# B&R Automation Studio project lab2_2 (part 2)

#### gmcipesm.cnc
```
Root (LangModule=ailgcode, Version=1.0)
  AILHeader = def ip_global BOOL  __CANCEL_RND 
    def ip_global BOOL  __C2_SPLINE_ACTIVE 
    def ip_global LREAL __RNDM_RADIUS 
    def ip_global LREAL __CSPLINE_CHORD_ERROR 
    def ip_global DINT __SET_GXX_ACTIVE 
    def ip_global DINT __SET_GXX_REACTIVATE 
    def ip_global DINT __SET_GXX_CALL_CNT 
    def ip_global REAL __VAR1 
    def ip_global DINT __ACTIVE_MIRROR 

    sub OnProgStartPrivate
      %__CANCEL_RND = 0;
      %__RNDM_RADIUS = 0.0;
      %__C2_SPLINE_ACTIVE = 0;
      %__CSPLINE_CHORD_ERROR = 0.001;
      %__SET_GXX_ACTIVE = 0;
      %__SET_GXX_REACTIVATE = 0;
      %__SET_GXX_CALL_CNT = 0;
      %__ACTIVE_MIRROR = 20;
    endsub

    sub EndSplineSection
      
      if (%__C2_SPLINE_ACTIVE)
        `T:GCodes,G802`(:"bc_par":1 :);
        %__C2_SPLINE_ACTIVE = 0;
        
        DispatchMPList(::);
      endif
    endsub
    sub WriteZpTable
      
      #next_motion.Command = MPCMD_SET_ZP_TABLE;
      #next_motion.Data.SetZeroPtTable.ZpRecIdx = $[1];
      #next_motion.Data.SetZeroPtTable.ZpOffset[0] = $[2];
      #next_motion.Data.SetZeroPtTable.ZpOffset[1] = $[3];
      #next_motion.Data.SetZeroPtTable.ZpOffset[2] = $[4];
      PushPacket(::);
      DispatchMPList(::);
    endsub

    sub ReactivateGxx
      
      
      if (%__SET_GXX_CALL_CNT != 0)
          if (%__SET_GXX_REACTIVATE == 1)
            `T:GCodes,G54`(::);
             DispatchMPList(::);
             #sys_vars.ZP = %__SET_GXX_REACTIVATE;
          elif (%__SET_GXX_REACTIVATE == 2)
            `T:GCodes,G55`(::);
             DispatchMPList(::);
             #sys_vars.ZP = %__SET_GXX_REACTIVATE;
          elif (%__SET_GXX_REACTIVATE == 3)
            `T:GCodes,G56`(::);
             DispatchMPList(::);
             #sys_vars.ZP = %__SET_GXX_REACTIVATE;
          elif (%__SET_GXX_REACTIVATE == 4)
            `T:GCodes,G57`(::);
             DispatchMPList(::);
             #sys_vars.ZP = %__SET_GXX_REACTIVATE;
          elif (%__SET_GXX_REACTIVATE == 5)
            `T:GCodes,G58`(::);
             DispatchMPList(::);
             #sys_vars.ZP = %__SET_GXX_REACTIVATE;
          elif (%__SET_GXX_REACTIVATE == 6)
            `T:GCodes,G59`(::);
             DispatchMPList(::);
             #sys_vars.ZP = %__SET_GXX_REACTIVATE;
          endif
          %__SET_GXX_REACTIVATE = 0;
          %__SET_GXX_CALL_CNT = 0;
      endif
    endsub (Append=Yes)
  BuiltInProcs:
    RESET_G54 = WriteZpTable(:1, 0.0, 0.0, 0.0:); (MinArgs=0, MaxArgs=0)
    RESET_G55 = WriteZpTable(:2, 0.0, 0.0, 0.0:); (MinArgs=0, MaxArgs=0)
    RESET_G56 = WriteZpTable(:3, 0.0, 0.0, 0.0:); (MinArgs=0, MaxArgs=0)
    RESET_G57 = WriteZpTable(:4, 0.0, 0.0, 0.0:); (MinArgs=0, MaxArgs=0)
    RESET_G58 = WriteZpTable(:5, 0.0, 0.0, 0.0:); (MinArgs=0, MaxArgs=0)
    RESET_G59 = WriteZpTable(:6, 0.0, 0.0, 0.0:); (MinArgs=0, MaxArgs=0)
    SET_G54 = WriteZpTable(:1, $[1], $[2], $[3]:);
      %_CNC.move_cmd_mode = MPCMD_LIN_INTPOL;
      %__SET_GXX_ACTIVE = 1;
      %__SET_GXX_REACTIVATE = 0;
      %__SET_GXX_CALL_CNT = 0;		
      
      `T:GCodes,G54`(::);
      #sys_vars.ZP = 1; (MinArgs=3, MaxArgs=3)
    SET_G55 = WriteZpTable(:2, $[1], $[2], $[3]:);
      %_CNC.move_cmd_mode = MPCMD_LIN_INTPOL;
      %__SET_GXX_ACTIVE = 2;
      %__SET_GXX_REACTIVATE = 0;
      %__SET_GXX_CALL_CNT = 0;		
      `T:GCodes,G55`(::);
      #sys_vars.ZP = 2; (MinArgs=3, MaxArgs=3)
    SET_G56 = WriteZpTable(:3, $[1], $[2], $[3]:);
      %_CNC.move_cmd_mode = MPCMD_LIN_INTPOL;
      %__SET_GXX_ACTIVE = 3;
      %__SET_GXX_REACTIVATE = 0;
      %__SET_GXX_CALL_CNT = 0;		
      `T:GCodes,G56`(::);
      #sys_vars.ZP = 3; (MinArgs=3, MaxArgs=3)
    SET_G57 = WriteZpTable(:4, $[1], $[2], $[3]:);
      %_CNC.move_cmd_mode = MPCMD_LIN_INTPOL;
      %__SET_GXX_ACTIVE = 4;
      %__SET_GXX_REACTIVATE = 0;
      %__SET_GXX_CALL_CNT = 0;		
      `T:GCodes,G57`(::);
      #sys_vars.ZP = 4; (MinArgs=3, MaxArgs=3)
    SET_G58 = WriteZpTable(:5, $[1], $[2], $[3]:);
      %_CNC.move_cmd_mode = MPCMD_LIN_INTPOL;
      %__SET_GXX_ACTIVE = 5;
      %__SET_GXX_REACTIVATE = 0;
      %__SET_GXX_CALL_CNT = 0;		
      `T:GCodes,G58`(::);
      #sys_vars.ZP = 5; (MinArgs=3, MaxArgs=3)
    SET_G59 = WriteZpTable(:6, $[1], $[2], $[3]:);
      %_CNC.move_cmd_mode = MPCMD_LIN_INTPOL;
      %__SET_GXX_ACTIVE = 6;
      %__SET_GXX_REACTIVATE = 0;
      %__SET_GXX_CALL_CNT = 0;		
      `T:GCodes,G59`(::);
      #sys_vars.ZP = 6; (MinArgs=3, MaxArgs=3)
    RESET_MIRROR = `T:GCodes,G20`(::); (MinArgs=0, MaxArgs=0)
  PVMacros:
    WORKFRAME $WFRAME (ArrayDims=0)
      SET = `T:BuiltInProcs,RESET_SCALING`(::);
        #next_motion.Data.Frame.Data = ${EXPR};
        #next_motion.Command = MPCMD_W_FRAME;
        PushPacket(::); (Inline=Yes)
    WORKFRAME_ADD $WFRAME_ADD (ArrayDims=0)
      SET = `T:BuiltInProcs,RESET_SCALING`(::);
        #next_motion.Data.Frame.Data = ${EXPR};
        #next_motion.Command = MPCMD_W_FRAME_ADD;
        PushPacket(::); (Inline=Yes)
  GCodes:
    G_INIT_ESM = ReactivateGxx(::); (GNum=-5, AutoPush=Yes, Eval=First, Inline=No, GenerateIfGroups=1,1000)
    G_MODAL (GNum=-1, AutoPush=Yes, Group=1000, Eval=Normal, IgnoreIfNoArgs=Yes)
      Arg (ref=dest, MinCount=0, MaxCount=NumAxes, NameType=AXISREF, DataType=PositionValue, WriteOpts=#:u?)
      Arg (ref=center, MinCount=0, MaxCount=3, NameType=InterpolParam, DataType=PositionValue, WriteOpts=#:u?)
      Arg (ref=circlept, MinCount=0, MaxCount=3, NameType=CirclePointParam, DataType=PositionValue, WriteOpts=#:u?)
      Arg (ref=angle, MinCount=0, MaxCount=1, NameType=RotationAngleSpecifier, DataType=RotationAngle, WriteOpts=#:u?)
      Arg (ref=radius, MinCount=0, MaxCount=1, NameType=RadiusSpecifier, DataType=RadiusValue, WriteOpts=#:u?)
    G00 = %_CNC.move_cmd_mode = MPCMD_RAPID_MOVE_INTPOL;
      #sys_vars.modal_grp1_set = 1;
      EndSplineSection(::); (GNum=0, Group=1,50, Inline=Yes, Eval=Early)
    G01 = %_CNC.move_cmd_mode = MPCMD_LIN_INTPOL;
      #sys_vars.modal_grp1_set = 1;
      EndSplineSection(::); (GNum=1, Group=1,50, Inline=Yes, Eval=Early)
    G02 = %_CNC.move_cmd_mode = MPCMD_CIRC_INTPOL_CW;
      #sys_vars.modal_grp1_set = 1;
      EndSplineSection(::); (GNum=2, Group=1,51, Inline=Yes, Eval=Early)
    G03 = %_CNC.move_cmd_mode = MPCMD_CIRC_INTPOL_CCW;
      #sys_vars.modal_grp1_set = 1;
      EndSplineSection(::); (GNum=3, Group=1,51, Inline=Yes, Eval=Early)
    G20 = #next_motion.Command = MPCMD_MIRRORING;
      #next_motion.Data.I4_value = 20;
      %__ACTIVE_MIRROR = #next_motion.Data.I4_value;
      PushPacket(::); (GNum=20, Group=3)
    G20.1 (GNum=20.1, Alias=MIRROR, Group=3)
      Arg (DataType=AXISREF, ref=axis1, MinCount=0, MaxCount=1)
      Arg (DataType=EqString, ref=eq, MinCount=0, MaxCount=1)
      Arg (DataType=FLOAT, ref=dummy_pos1, MinCount=0, MaxCount=1)
      Arg (DataType=AXISREF, ref=axis2, MinCount=0, MaxCount=1)
      Arg (DataType=EqString, ref=eq, MinCount=0, MaxCount=1)
      Arg (DataType=FLOAT, ref=dummy_pos2, MinCount=0, MaxCount=1)
    G20.2 (GNum=20.2, Alias=AMIRROR, Group=3)
      Arg (DataType=AXISREF, ref=axis1, MinCount=1, MaxCount=1)
      Arg (DataType=EqString, ref=eq, MinCount=0, MaxCount=1)
      Arg (DataType=FLOAT, ref=dummy_pos1, MinCount=0, MaxCount=1)
      Arg (DataType=AXISREF, ref=axis2, MinCount=0, MaxCount=1)
      Arg (DataType=EqString, ref=eq, MinCount=0, MaxCount=1)
      Arg (DataType=FLOAT, ref=dummy_pos2, MinCount=0, MaxCount=1)
    G21 = #next_motion.Command = MPCMD_MIRRORING;
      #next_motion.Data.I4_value = 21;
      %__ACTIVE_MIRROR = #next_motion.Data.I4_value;
      PushPacket(::); (GNum=21, Group=3)
    G22 = #next_motion.Command = MPCMD_MIRRORING;
      #next_motion.Data.I4_value = 22;
      %__ACTIVE_MIRROR = #next_motion.Data.I4_value;
      PushPacket(::); (GNum=22, Group=3)
    G23 = #next_motion.Command = MPCMD_MIRRORING;
      #next_motion.Data.I4_value = 23;
      %__ACTIVE_MIRROR = #next_motion.Data.I4_value;
      PushPacket(::); (GNum=23, Group=3)
    G25.1 (GNum=25.1, Group=11, Alias=RNDM)
      Arg (NameType=EqString, DataType=TangArcRadius, ref=radius)
    G25.2 (GNum=25.2, Group=11, Alias=RND)
      Arg (NameType=EqString, DataType=TangArcRadius, ref=radius)
    G53 = #next_motion.Command = MPCMD_ABS_ZP_SHIFT;
      #next_motion.Data.AbsZeroPtShift.ZpRecIdx = 0;
      PushPacket(::);
      #sys_vars.ZP = 0;
      
      %__SET_GXX_REACTIVATE = %__SET_GXX_ACTIVE;
      %__SET_GXX_CALL_CNT = 0; (GNum=53, Group=6, AllowGroups=8,19,21,100,101,102,103)
    G92 (GNum=92, Group=21, ResetArgs=Yes, AllowGroups=6,8,19,32,100,101,102,103)
      Arg (NameType=AXISREF, DataType=PositionValue, ref=offset, MinCount=0, MaxCount=NumAxes, WriteOpts=#:u?)
      Arg (NameType=RotationAngleSpecifier, DataType=RotationAngle, ref=h_rot, MinCount=0, MaxCount=1, WriteOpts=#:u?, DenyArgs=3,4,5)
      Arg (NameType=EulerAngleName, DataType=RotationAngle, ref=e_rot, MinCount=0, MaxCount=3, WriteOpts=#:u?, DenyArgs=2,4,5)
      Arg (NameType=RPYAngleName, DataType=RotationAngle, ref=rpy_rot, MinCount=0, MaxCount=3, WriteOpts=#:u?, DenyArgs=2,3,5)
      Arg (NameType=RotaryVectorName, DataType=RotaryVector, ref=matrix, MinCount=0, MaxCount=3, WriteOpts=#:u?, DenyArgs=2,3,4)
    G92.1 (GNum=92.1, Group=21, ALIAS=SCALE, AliasIsPattern=Yes)
      Arg (DataType=FLOAT, ref=factor, MinCount=0, MaxCount=1)
    G92.2 (GNum=92.2, Group=21, ALIAS=ASCALE, AliasIsPattern=Yes)
      Arg (DataType=FLOAT, ref=factor, MinCount=1, MaxCount=1)
    G492 (GNum=492, Group=490, Alias=TRANS, AllowGroups=9999)
      Arg (NameType=AXISREF, DataType=PositionValue, ref=offsets, MinCount=0, MaxCount=NumAxes, WriteOpts=#:)
    G494 (GNum=494, Group=490, Alias=ROT, AllowGroups=9999, MinArgs=0, MaxArgs=1)
      Arg RPLArgPrefix (DataType=FLOAT, ref=rpl_value, MinCount=0, MaxCount=1, DenyArgs=offsets)
      Arg (NameType=AXISREF, DataType=PositionValue, ref=offsets, MinCount=0, MaxCount=NumAxes, DenyArgs=rpl_value, WriteOpts=#:)
    G500 = %__SET_GXX_REACTIVATE = 0;
       %__SET_GXX_ACTIVE = 0;
       %__SET_GXX_CALL_CNT = 0;
      `T:GCodes,G53`(::); (GNum=500, Group=6, AllowGroups=8,19,21,100,101,102,103)
    G804 = if (!%__C2_SPLINE_ACTIVE)
         
        `T:GCodes,G801`(:"seg_type":"CE", "seg_par":%__CSPLINE_CHORD_ERROR, "bc_par":1 :);
        %__C2_SPLINE_ACTIVE = 1;
        
        DispatchMPList(::);
        
        %_CNC.move_cmd_mode = MPCMD_LIN_INTPOL;
      endif (GNum=804, Alias=CSPLINE)
```

### Data object Logical/GmcIpConfig/gmcipmxd (Cnc, version 5.02.1)

#### gmcipmxd.cnc
```
(********************************************************************
 * COPYRIGHT (C) B&R Industrial Automation GmbH
 ********************************************************************
 * Library: Motion Command Extension
 * File: arnc0mx.typ
 * Author: B&R
 ********************************************************************
 * Data types of Motion Command Library
 ********************************************************************)

TYPE
	MXOrientationType : STRUCT
		Type : UDINT;
		Angle : ARRAY[0..3]OF LREAL;
	END_STRUCT;
	MXPositionType : STRUCT
		x : LREAL;
		y : LREAL;
		z : LREAL;
	END_STRUCT;
	MXFrameType : 	STRUCT
		Pos : MXPositionType;
		Orient : MXOrientationType;
	END_STRUCT;
	MXToolType : STRUCT
		Index : UDINT;
		Frame : MXFrameType;
		Radius : LREAL;
	END_STRUCT;
	MXJointAxisType :ARRAY[0..5]OF LREAL;
	MXAuxAxisType :ARRAY[0..14]OF LREAL;
	MXBaseAxisType :ARRAY[0..5]OF LREAL;
	MXRotAxisType :ARRAY[0..5]OF LREAL;
	MXConfigType : 	STRUCT
		Mode : UDINT;
	END_STRUCT;
	MXPointType : 	STRUCT
		Pos : MXPositionType;
		Orient : MXOrientationType;
		Cfg : MXConfigType;
		RotAxis : MXRotAxisType;
		AuxAxis : MXAuxAxisType;
	END_STRUCT;
	MXPathTransType : STRUCT
		Radius	:	LREAL;
		Type	:	UDINT;
	END_STRUCT;
	MXPathDescType : STRUCT
		Trans	:	MXPathTransType;
	END_STRUCT;
	MXOptMotType : STRUCT
		Enable : BOOL;
		VelPathDef : USINT;
		RobotPar : USINT;
		Limits : USINT;
	END_STRUCT;
	MXDynamicDescType :	STRUCT
		Accel : LREAL := 100;
		Decel : LREAL := 100;
		Optmot : MXOptMotType;
	END_STRUCT;
	MXHWTrigType : 	STRUCT
		Source : USINT;
		Index : USINT;
	END_STRUCT;
	MXSWTrigType : STRUCT
		Expression : STRING[64];
	END_STRUCT;
	MXTriggConfigType :	STRUCT
		Type : UINT;
		HWTrig : MXHWTrigType;
		SWTrig : MXSWTrigType;
		Edge : USINT;
		ResidPath : USINT;
	END_STRUCT;
	MXVelocityType : STRUCT
		v : LREAL;
		Mode : UDINT := 1;
	END_STRUCT;
	MXAxisTargetType : 	STRUCT
		JointAxis : MXJointAxisType;
		AuxAxis : MXAuxAxisType;
		BaseAxis : MXBaseAxisType;
	END_STRUCT;
	MXCDCType : STRUCT
		ArcTransSpd : LREAL := 100;
		SpdMode : UDINT;
		ContourViolation : UDINT;
		TransMode : UDINT;
		EntryMode : USINT;
		AcrToLine : BOOL;
	END_STRUCT;
	MXAutoTangType : STRUCT
		Offset : LREAL;
	END_STRUCT;
	MXHWTriggerType :	STRUCT
		Source : UINT;
		Index : UINT;
	END_STRUCT;
	MXTriggerConfigType : 	STRUCT
		Type : UINT;
		Edge : UINT;
		HWTrigger : MXHWTriggerType;
	END_STRUCT;
END_TYPE

(********************************************************************
 * COPYRIGHT (C) B&R Industrial Automation GmbH
 ********************************************************************
 * Library: ARNC0MX
 * File: arnc0mx.fun
 * Created: 13.06.2012
 ********************************************************************
 * Functions and function blocks of library ARNC0MX
 ********************************************************************)
FUNCTION MXPointToJointEx1 : UDINT
	VAR_INPUT
		AddrTrfData : UDINT;
		Point : MXPointType;
		Joint : MXJointAxisType;
		TrfType : UDINT;
		Tool : MXToolType;
		BaseFrame : MXFrameType;
		RefJoint : ARRAY[0..5] OF LREAL;
	END_VAR
END_FUNCTION

FUNCTION MXPointToJointEx : UDINT
	VAR_INPUT
		AddrTrfData : UDINT;
		Point : MXPointType;
		Joint : MXJointAxisType;
		TrfType : UDINT;
		Tool : MXToolType;
		BaseFrame : MXFrameType;
		RefJoint : MXJointAxisType;
	END_VAR
END_FUNCTION

FUNCTION MXJointToPointEx1 : UDINT
	VAR_INPUT
		AddrTrfData : UDINT;
		Joint : MXJointAxisType;
		Point : MXPointType;
		AnglesType : UDINT;
		TrfType : UDINT;
		Tool : MXToolType;
		BaseFrame : MXFrameType;
		RefPath : ARRAY[0..5] OF LREAL;
	END_VAR
END_FUNCTION

FUNCTION MXJointToPointEx : UDINT
	VAR_INPUT
		AddrTrfData : UDINT;
		Joint : MXJointAxisType;
		Point : MXPointType;
		AnglesType : UDINT;
		TrfType : UDINT;
		Tool : MXToolType;
		BaseFrame : MXFrameType;
		RefPoint : MXPointType;
	END_VAR
END_FUNCTION

FUNCTION MXCncAxesToPoint : UDINT
	VAR_INPUT
		AddrTrfData : UDINT;
		Axis : ARRAY[0..14] OF LREAL;
		Point : MXPointType;
		TrfType : UDINT;
		AnglesType : UDINT;
		AxisMapCode : ARRAY[0..14] OF UINT;
		AxisMapIdx : ARRAY[0..14] OF UINT;
		ActiveAxesCount : UDINT;
	END_VAR
END_FUNCTION

FUNCTION MXFromOrient : UDINT
	VAR_INPUT
		Orient : MXOrientationType;
		Matrix : ARRAY[0..8] OF LREAL;
	END_VAR
END_FUNCTION

FUNCTION MXToOrient : UDINT
	VAR_INPUT
		Matrix : ARRAY[0..8] OF LREAL;
		Type : UDINT;
		Orient : MXOrientationType;
		RefAngle : ARRAY[0..2] OF LREAL;
	END_VAR
END_FUNCTION

FUNCTION MXConvertOrient : UDINT
	VAR_INPUT
		OrientIn : MXOrientationType;
		Type : UDINT;
		OrientOut : MXOrientationType;
		RefAngle : ARRAY[0..2] OF LREAL;
	END_VAR
END_FUNCTION

FUNCTION MXFrameRotX : UDINT
	VAR_INPUT
		Frame : MXFrameType;
		Angle : LREAL;
	END_VAR
END_FUNCTION

FUNCTION MXFrameRotY : UDINT
	VAR_INPUT
		Frame : MXFrameType;
		Angle : LREAL;
	END_VAR
END_FUNCTION

FUNCTION MXFrameRotZ : UDINT
	VAR_INPUT
		Frame : MXFrameType;
		Angle : LREAL;
	END_VAR
END_FUNCTION

FUNCTION MXFrameEuler : UDINT
	VAR_INPUT
		Frame : MXFrameType;
		Phi : LREAL;
		Theta : LREAL;
		Psi : LREAL;
	END_VAR
END_FUNCTION

FUNCTION MXFrameRPY : UDINT
	VAR_INPUT
		Frame : MXFrameType;
		Roll : LREAL;
		Pitch : LREAL;
		Yaw : LREAL;
	END_VAR
END_FUNCTION

FUNCTION MXFrameTrans : UDINT
	VAR_INPUT
		Frame : MXFrameType;
		DistanceX : LREAL;
		DistanceY : LREAL;
		DistanceZ : LREAL;
	END_VAR
END_FUNCTION

FUNCTION MXFrameTransX : UDINT
	VAR_INPUT
		Frame : MXFrameType;
		Distance : LREAL;
	END_VAR
END_FUNCTION

FUNCTION MXFrameTransY : UDINT
	VAR_INPUT
		Frame : MXFrameType;
		Distance : LREAL;
	END_VAR
END_FUNCTION

FUNCTION MXFrameTransZ : UDINT
	VAR_INPUT
		Frame : MXFrameType;
		Distance : LREAL;
	END_VAR
END_FUNCTION

FUNCTION MXFrameApply : UDINT
	VAR_INPUT
		Frame1 : MXFrameType;
		Frame2 : MXFrameType;
	END_VAR
END_FUNCTION

FUNCTION MXFromFrame : UDINT
	VAR_INPUT
		Frame : MXFrameType;
		PointIn : MXPointType;
		PointOut : MXPointType;
	END_VAR
END_FUNCTION

FUNCTION MXToFrame : UDINT
	VAR_INPUT
		Frame : MXFrameType;
		PointIn : MXPointType;
		PointOut : MXPointType;
	END_VAR
END_FUNCTION

(********************************************************************
 * COPYRIGHT (C) B&R Industrial Automation GmbH
 ********************************************************************
 * Library: Motion Command Extension
 * File: arnc0mx.var
 * Author: B&R
 ********************************************************************
 * Constants of Motion Command Library
 ********************************************************************)

(* Velocity mode constants (<MXVelocityType>.Mode) *)
VAR CONSTANT
  MX_VEL_MODE_RAPID : UDINT := 0; (* rapid mode *)
  MX_VEL_MODE_FEED  : UDINT := 1; (* feedrate mode *)
  MX_VEL_MODE_TIME  : UDINT := 2; (* inverse time mode *)
END_VAR

(* MXVelocityType constants *)
VAR CONSTANT
  MX_VEL_RAPID  : MXVelocityType := (Mode:=0);           (* rapid movement         *)
  MX_VEL_F50000 : MXVelocityType := (v:=50000, Mode:=1); (* 50000 units per minute *)
  MX_VEL_F10000 : MXVelocityType := (v:=10000, Mode:=1); (* 10000 units per minute *)
  MX_VEL_F5000  : MXVelocityType := (v:=5000,  Mode:=1); (* 5000 units per minute  *)
  MX_VEL_F1000  : MXVelocityType := (v:=1000,  Mode:=1); (* 1000 units per minute  *)
  MX_VEL_F500   : MXVelocityType := (v:=500,   Mode:=1); (* 500 units per minute   *)
  MX_VEL_F100   : MXVelocityType := (v:=100,   Mode:=1); (* 100 units per minute   *)
END_VAR

(* Trigger configuration constants *)
VAR CONSTANT
  MX_TRIGGER_HW	            : UINT := 0;           (* Hardware trigger - MXHWTriggerType *)
  MX_TRIGGER_POSITIVE_EDGE  : UINT := 0;           (* Positive edge						 *)
  MX_TRIGGER_NEGATIVE_EDGE  : UINT := 1;           (* Negative edge						 *)
  MX_TRIGGER_HW_INPUT1		: UINT := 1;           (* Hardware trigger input 1			 *)
  MX_TRIGGER_HW_INPUT2		: UINT := 2;           (* Hardware trigger input 1			 *)
END_VAR

(* MXFrameMXFrameType constants *)
VAR CONSTANT
  MX_FRM_ZERO : MXFrameType := (0); (* zero (identity) frame *)
END_VAR

(* Transition type constants (<MXPathTransType>.Type) *)
VAR CONSTANT
  MX_TRANS_OFF      : UDINT := 0; (* Transition deactivated *)
  MX_TRANS_ACCURATE : UDINT := 1; (* Accuracy hold *)
  MX_TRANS_ARC      : UDINT := 2; (* Tangential transition arcs *)
  MX_TRANS_ROUND    : UDINT := 3; (* Rounding edges *)
END_VAR

(* Orientation type constants (<MXOrientationType>.Type) matches constants from TRF_LIB *)
VAR CONSTANT
  MX_CARDAN_XYZ_ANGLES    : UDINT := 1;      (* Cardan XYZ angles *)
  MX_EULER_XYZ_ANGLES     : UDINT := 1;      (* Cardan XYZ angles *)
  MX_CARDAN_XZY_ANGLES    : UDINT := 2;      (* Cardan XZY angles *)
  MX_EULER_XZY_ANGLES     : UDINT := 2;      (* Cardan XZY angles *)
  MX_CARDAN_YXZ_ANGLES    : UDINT := 4;      (* Cardan YXZ angles *)
  MX_EULER_YXZ_ANGLES     : UDINT := 4;      (* Cardan YXZ angles *)
  MX_CARDAN_YZX_ANGLES    : UDINT := 8;      (* Cardan YZX angles *)
  MX_EULER_YZX_ANGLES     : UDINT := 8;      (* Cardan YZX angles *)
  MX_CARDAN_ZXY_ANGLES    : UDINT := 16;     (* Cardan ZXY angles *)
  MX_EULER_ZXY_ANGLES     : UDINT := 16;     (* Cardan ZXY angles *)
  MX_CARDAN_ZYX_ANGLES    : UDINT := 32;     (* Cardan ZYX angles *)
  MX_EULER_ZYX_ANGLES     : UDINT := 32;     (* Cardan ZYX angles *)
  MX_EULER_XYX_ANGLES     : UDINT := 64;     (* Euler XYX angles  *)
  MX_EULER_XZX_ANGLES     : UDINT := 128;    (* Euler XZX angles  *)
  MX_EULER_YXY_ANGLES     : UDINT := 256;    (* Euler YXY angles  *)
  MX_EULER_YZY_ANGLES     : UDINT := 512;    (* Euler YZY angles  *)
  MX_EULER_ZXZ_ANGLES     : UDINT := 1024;   (* Euler ZXZ angles  *)
  MX_EULER_ZYZ_ANGLES     : UDINT := 2048;   (* Euler ZYZ angles  *)
  MX_POSITIVE_ANGLES      : UDINT := 4096;   (* mathematically positive angles *)
  MX_NEGATIVE_ANGLES      : UDINT := 8192;   (* mathematically negative angles *)
  MX_DIRECT_ANGLES        : UDINT := 16384;  (* direct "R" rotation matrix     *)
  MX_INDIRECT_ANGLES      : UDINT := 32768;  (* indirect "R^T" rotation matrix *)
  MX_EULER_ANGLES         : UDINT := 1024;   (* Euler ZXZ is commonly in view  *)
  MX_CARDAN_ANGLES        : UDINT := 1;      (* Cardan XYZ is commonly in view *)
  MX_NAUTICAL_ANGLES      : UDINT := 1;      (* Cardan XYZ is commonly in view *)
  MX_TAIT_BRYAN_ANGLES    : UDINT := 1;      (* Cardan XYZ is commonly in view *)
  MX_QUATERNION           : UDINT := 8000;   (* quaternion *)
END_VAR

(* Kinematics configuration mode constants (<MXConfigType>.Mode) matches constants from TRF_LIB *)
VAR CONSTANT
  MX_MODE_FRONT           : UDINT := 1;          (* front *)
  MX_MODE_BACK            : UDINT := 2;          (* back *)
  MX_MODE_CONVEX          : UDINT := 4;          (* convex *)
  MX_MODE_CONCAVE         : UDINT := 8;          (* concave *)
  MX_MODE_POSITIVE        : UDINT := 16;         (* positive *)
  MX_MODE_NEGATIVE        : UDINT := 32;         (* negative *)
  MX_MODE_LEFT            : UDINT := 64;         (* left *)
  MX_MODE_RIGHT           : UDINT := 128;        (* right *)
  MX_MODE_DIRECT          : UDINT := 256;        (* direct *)
  MX_MODE_INDIRECT        : UDINT := 512;        (* indirect *)
  MX_MODE_CONVEX2         : UDINT := 1024;       (* convex2 *)
  MX_MODE_CONCAVE2        : UDINT := 2048;       (* concave2 *)
  MX_MODE_CONVEX3         : UDINT := 4096;       (* convex3 *)
  MX_MODE_CONCAVE3        : UDINT := 8192;       (* concave3 *)
  MX_MODE_HETEROGENEOUS   : UDINT := 16384;      (* heterogeneous *)
  MX_MODE_HOMOGENEOUS     : UDINT := 32768;      (* homogeneous *)
  MX_MODE_LEFT2           : UDINT := 65536;      (* left2 *)
  MX_MODE_RIGHT2          : UDINT := 131072;     (* right2 *)
  MX_MODE_NEG_DIR         : UDINT := 268435456;  (* negative direction forced *)
  MX_MODE_POS_DIR         : UDINT := 536870912;  (* positive direction forced *)
  MX_MODE_IN_SW_ENDS      : UDINT := 1073741824; (* in SW ends *)
END_VAR

(* Cutter diameter compensation constants *)
VAR CONSTANT
  MX_CDC_LEFT                    : UDINT := 0;      (* CDC left *)
  MX_CDC_RIGHT                   : UDINT := 1;      (* CDC right *)
  MX_CDC_SPD_ON_CONTOUR          : UDINT := 0;      (* Path speed moves to the contour *)
  MX_CDC_SPD_ON_TCP              : UDINT := 1;      (* Path speed moves to the center of the tool *)
  MX_CDC_NO_COUNTER_VIOLATION    : UDINT := 0;      (* Do NOT allow contour violations due to very short path *)
  MX_CDC_VIOLATION_SHORT_PATH    : UDINT := 1;      (* Allow contour violations due to very short path sections *)
  MX_CDC_VIOLATION_INNER_EDGE    : UDINT := 2;      (* Allow contour violations due to an inner edge without intersection *)
  MX_CDC_LINEAR_TRANSITION       : UDINT := 0;      (* CDC with linear transitions *)
  MX_CDC_ARC_TRANSITION          : UDINT := 1;      (* CDC with arc transitions *)
  MX_CDC_ENTRY_BLOCK             : UDINT := 0;      (* Activate/deactivate CDC indirectly with transi-tion block *)
  MX_CDC_ENTRY_DIRECT            : UDINT := 1;      (* Activate/deactivate CDC directly *)
  MX_CDC_ENTRY_INDIRECT          : UDINT := 2;      (* Activate/deactivate CDC indirectly *)
  MX_CDC_NO_ARC_TO_LINE          : UDINT := 0;      (* Deactivate replacement of arc with straight line *)
  MX_CDC_ARC_TO_LINE             : UDINT := 1;      (* Activate replacement of arc with straight line *)
END_VAR

(* Transformation function types *)
VAR CONSTANT
  MX_TRF_TYPE_INVERSE            : UDINT := 0;      (* TRF_inverse  function *)
  MX_TRF_TYPE_INVERSE2           : UDINT := 1;      (* TRF_inverse2 function *)
  MX_TRF_TYPE_INVERSE3           : UDINT := 2;      (* TRF_inverse3 function *)
  MX_TRF_TYPE_DIRECT             : UDINT := 0;      (* TRF_direct   function *)
  MX_TRF_TYPE_DIRECT2            : UDINT := 1;      (* TRF_direct2  function *)
  MX_TRF_TYPE_DIRECT3            : UDINT := 2;      (* TRF_direct3  function *)
END_VAR

(* Statuses, warnings, errors *)
VAR CONSTANT
  MX_OK                          : UDINT := 0;     (* Status OK *)
  MX_WARNING_AXES                : UDINT := 2001;  (* Transformation returns valid values with warnings on axes *)
  MX_WARNING_REF_POINT_ANGLES    : UDINT := 2002;  (* Values in reference point or reference joint axes may be ignored due to conversion to another angles type *)
  MX_ERROR_WRONG_ANGLE_TYPE      : UDINT := 6001;  (* Angles type is not supported *)
  MX_ERROR_TRF_DATA_NOT_DEFINED  : UDINT := 6002;  (* Address of the transformation data variable is zero *)
  MX_ERROR_WRONG_ROBOT           : UDINT := 6003;  (* Robot is not supported *)
  MX_ERROR_WRONG_TRF_TYPE        : UDINT := 6004;  (* Transformation type not supported *)
  MX_ERROR_TRF_LIB_NOT_SUPPORTED : UDINT := 6005;  (* Transformation library of not supported version *)
  MX_ERROR_TRF_CMD_CODE			 : UDINT := 8001;  (* Unknown command code *)
  MX_ERROR_TRF_MEASURE           : UDINT := 8002;  (* Unknown measure *)
  MX_ERROR_TRF_ANGLES_TYPE       : UDINT := 8003;  (* Unknown angles type *)
  MX_ERROR_TRF_GEN29_CMD_CODE    : UDINT := 9001;  (* Unknown command code *)
  MX_ERROR_UNKNOWN_ROBOT         : UDINT := 9002;  (* Unknown robot *)
  MX_ERROR_INVALID_TRF_TYPE      : UDINT := 9003;  (* Invalid type of transformation *)
  MX_ERROR_TRF_ERROR_AXES        : UDINT := 10003; (* Transformation function returns error of axis *)
  MX_ERROR_TRF_NOT_LICENSED      : UDINT := 10008; (* Transformation function not licenced *)
  MX_ERROR_TRF_NOT_SUPPORTED     : UDINT := 10009; (* Transformation function not supported *)
  MX_ERROR_FCT_NOT_DEFINED       : UDINT := 10010; (* Transformation function address is zero *)
  MX_ERROR_TRF_INVALID_INPUTS    : UDINT := 10015; (* Invalid inputs for transformation error *)
END_VAR

(* Error offsets *)
VAR CONSTANT
  MX_OFFSET_WARNING              : UDINT := 2000;  (* ARNC0MX warnings *)
  MX_OFFSET_WARNING_TRF_FUN      : UDINT := 4000;  (* TRF_LIB warnings *)
  MX_OFFSET_ERROR                : UDINT := 6000;  (* ARNC0MX errros *)
  MX_OFFSET_ERROR_TRF_FUN        : UDINT := 12000; (* TRF_LIB errors *)
END_VAR

(********************************************************************
 * COPYRIGHT (C) B&R Industrial Automation GmbH
 ********************************************************************
 * Library: Motion Command Library
 * File: arnc0mxsv.var
 * Author: B&R
 ********************************************************************
 * System Variables of Motion Command Library
 ********************************************************************)
VAR {SHARED_IP_GLOBAL}
   _Frm  : MXFrameType;
   _Tool : MXToolType;
   _Vel  : MXVelocityType;
   _Base : MXFrameType;
   _Ref  : MXJointAxisType;
   _Pth  : MXPathDescType;
   _Dyn  : MXDynamicDescType;
END_VAR

VAR CONSTANT
   FRM_0   : MXFrameType := (0);
   POINT_0 : MXPointType := (0);
   BASE_0  : MXFrameType := (0);
   TOOL_0  : MXToolType  := (0);
   VEL_0   : MXVelocityType := (Mode:=1);
   REF_0   : MXJointAxisType := (0);
   VEC6_0  : ARRAY[0..5] OF LREAL := 6(0.0);
   PTH_0   : MXPathDescType := (0);
   DYN_0   : MXDynamicDescType := (Accel:=100, Decel:=100);
   AXIS_TARGET_0 : MXAxisTargetType := (0);
END_VAR

VAR {SHARED_IP_GLOBAL}
  __tmp_point : MXPointType;
  __tmp_frame : MXFrameType;
  __tmp_tool : MXToolType;
  __tmp_vel : MXVelocityType;
  __tmp_joint_axis : MXJointAxisType;
  __tmp_axis_target : MXAxisTargetType;
  __tmp_pth : MXPathDescType;
  __tmp_dynamic : MXDynamicDescType;
  __tmp_cdc : MXCDCType;
  __tmp_auto_tang : MXAutoTangType;
  __tmp_trigger : MXTriggerConfigType;
  __mx_status : UDINT;
  __tmp_vec6 : ARRAY[0..5] OF LREAL;
  __tmp_set_pos : ARRAY[0..14] OF LREAL;
  __tmp_axis_code : ARRAY[0..14] OF UINT;
  __tmp_axis_idx : ARRAY[0..14] OF UINT;
END_VAR
```

### Data object Logical/GmcIpConfig/gmcipmx (Cnc, version 5.02.1)

#### gmcipmx.cnc
```
Root (LangModule=ailgcode, Version=1.0)
  AILHeader = sub OnProgStartPrivate
      %_Frm = %FRM_0;
      %_Base = %BASE_0;
      %_Tool = %TOOL_0;
      %_Vel = %VEL_0;
      %_Pth = %PTH_0;
      %_Dyn = %DYN_0;
      if (%_CNC.optmot_segmentation_on)
        %_Dyn.Optmot.Enable = 1 
      endif      
      BlockCpy(:\%_Ref, \%REF_0:);
    endsub
  BuiltInProcs:
    WAIT_PP_SYNC = #next_motion.Command = MPCMD_IP_SYNCH_PP;
      PushPacket(::);
      DispatchAndWait(:IPCMD_SYNC_PP_CONT:);
    ERROR_EX = ErrorEx(:"id":$[1],"fmt":$[2],"data":(:$[3],$[4],$[5],$[6],$[7],$[8],$[9],$[10],$[11],$[12],$[13],$[14]:):); (MinArgs=3, MaxArgs=14)
    SET_POINT:
      Arg (ref=POINT, DataType=ANY_DATA, MinCount=1, MaxCount=1)
    SET_TRIGGER_CONFIG:
      Arg (ref=TRIGGER, DataType=ANY_DATA, MinCount=1, MaxCount=1)
      Arg (ref=bHALT, DataType=ANY_DATA, MinCount=1, MaxCount=1)
      Arg (ref=ID, DataType=ANY_DATA, MinCount=1, MaxCount=1)
    SET_WANTED_JOINT:
      Arg (ref=Ref, DataType=ANY_DATA, MinCount=1, MaxCount=1)
    SET_CIRCLE:
      Arg (ref=END_POINT, DataType=ANY_DATA, MinCount=1, MaxCount=1)
      Arg (ref=CIRCLE_POINT, DataType=ANY_DATA, MinCount=1, MaxCount=1)
      Arg (ref=Angle, DataType=IEC_LREAL, MinCount=0, MaxCount=1)
    SET_AXIS_TARGET:
      Arg (ref=AXIS_TARGET, DataType=ANY_DATA, MinCount=1, MaxCount=1)
    SET_FRAME:
      Arg (ref=Frm, DataType=ANY_DATA, MinCount=0, MaxCount=1)
    SET_BASEFRAME:
      Arg (ref=Base, DataType=ANY_DATA, MinCount=0, MaxCount=1)
    SET_TOOL:
      Arg (ref=Tool, DataType=ANY_DATA, MinCount=0, MaxCount=1)
    SET_PATH_DESC:
      Arg (ref=Pth, DataType=ANY_DATA, MinCount=0, MaxCount=1)
    SET_DYNAMIC_DESC:
      Arg (ref=Dyn, DataType=ANY_DATA, MinCount=0, MaxCount=1)
    SET_VELOCITY:
      Arg (ref=Vel, DataType=ANY_DATA, MinCount=0, MaxCount=1)
    JointToPoint:
      Arg (ref=Joint, UserType=MXJointAxisType, MinCount=1, MaxCount=1)
      Arg (ref=Point, UserType=MXPointType, MinCount=1, MaxCount=1)
    PointToJoint:
      Arg (ref=Point, UserType=MXPointType, MinCount=1, MaxCount=1)
      Arg (ref=Joint, UserType=MXJointAxisType, MinCount=1, MaxCount=1)
    MoveL:
      Arg (ref=POINT, UserType=MXPointType, MinCount=1, MaxCount=1)
      Arg (ref=Frm, UserType=MXFrameType, MinCount=0, MaxCount=1)
      Arg (ref=Base, UserType=MXFrameType, MinCount=0, MaxCount=1)
      Arg (ref=Tool, UserType=MXToolType, MinCount=0, MaxCount=1)
      Arg (ref=Vel, UserType=MXVelocityType, MinCount=0, MaxCount=1)
      Arg (ref=Pth, UserType=MXPathDescType, MinCount=0, MaxCount=1)
      Arg (ref=Dyn, UserType=MXDynamicDescType, MinCount=0, MaxCount=1)
    MoveJ:
      Arg (ref=POINT, UserType=MXPointType, MinCount=1, MaxCount=1)
      Arg (ref=Frm, UserType=MXFrameType, MinCount=0, MaxCount=1)
      Arg (ref=Base, UserType=MXFrameType, MinCount=0, MaxCount=1)
      Arg (ref=Tool, UserType=MXToolType, MinCount=0, MaxCount=1)
      Arg (ref=Vel, UserType=MXVelocityType, MinCount=0, MaxCount=1)
      Arg (ref=Ref, UserType=MXJointAxisType, MinCount=0, MaxCount=1)
      Arg (ref=Pth, UserType=MXPathDescType, MinCount=0, MaxCount=1)
      Arg (ref=Dyn, UserType=MXDynamicDescType, MinCount=0, MaxCount=1)
    MoveC:
      Arg (ref=END_POINT, UserType=MXPointType, MinCount=1, MaxCount=1)
      Arg (ref=CIRCLE_POINT, UserType=MXPointType, MinCount=1, MaxCount=1)
      Arg (ref=Angle, DataType=IEC_LREAL, MinCount=0, MaxCount=1)
      Arg (ref=Frm, UserType=MXFrameType, MinCount=0, MaxCount=1)
      Arg (ref=Base, UserType=MXFrameType, MinCount=0, MaxCount=1)
      Arg (ref=Tool, UserType=MXToolType, MinCount=0, MaxCount=1)
      Arg (ref=Vel, UserType=MXVelocityType, MinCount=0, MaxCount=1)
      Arg (ref=Pth, UserType=MXPathDescType, MinCount=0, MaxCount=1)
      Arg (ref=Dyn, UserType=MXDynamicDescType, MinCount=0, MaxCount=1)
    MoveA:
      Arg (ref=AXIS_TARGET, UserType=MXAxisTargetType, MinCount=1, MaxCount=1)
      Arg (ref=Vel, UserType=MXVelocityType, MinCount=0, MaxCount=1)
      Arg (ref=Dyn, UserType=MXDynamicDescType, MinCount=0, MaxCount=1)
      Arg (ref=Pth, UserType=MXPathDescType, MinCount=0, MaxCount=1)
    MoveLSearch:
      Arg (ref=POINT, UserType=MXPointType, MinCount=1, MaxCount=1)
      Arg (ref=TRIGGER, UserType=MXTriggerConfigType, MinCount=1, MaxCount=1)
      Arg (ref=bHALT, DataType=IEC_BOOL, MinCount=1, MaxCount=1)
      Arg (ref=ID, DataType=IEC_UINT, MinCount=1, MaxCount=1)
      Arg (ref=Frm, UserType=MXFrameType, MinCount=0, MaxCount=1)
      Arg (ref=Base, UserType=MXFrameType, MinCount=0, MaxCount=1)
      Arg (ref=Tool, UserType=MXToolType, MinCount=0, MaxCount=1)
      Arg (ref=Vel, UserType=MXVelocityType, MinCount=0, MaxCount=1)
      Arg (ref=Pth, UserType=MXPathDescType, MinCount=0, MaxCount=1)
      Arg (ref=Dyn, UserType=MXDynamicDescType, MinCount=0, MaxCount=1)
    WaitTime:
      Arg (ref=set_time, DataType=IEC_LREAL, MinCount=1, MaxCount=1)
    WaitIp = #next_motion.Command = MPCMD_IP_SYNCH;
      if (#thread.restart.playback)
        #next_motion.Data.I4_value = ncSIMULATION;
      else
        #next_motion.Data.I4_value = ncSTANDARD;
      endif
      PushPacket(::);
      DispatchAndWait(:IPCMD_SYNC_PLC_CONT:);
    WaitEndMove = #next_motion.Command = MPCMD_IP_SYNCH_PATH;
      PushPacket(::);
      DispatchAndWait(:IPCMD_SYNC_PATH_CONT:);
    TmpTool = %__tmp_tool.Frame.Pos.x = %_CNC.tool_dx;
      %__tmp_tool.Frame.Pos.y = %_CNC.tool_dy;
      %__tmp_tool.Frame.Pos.z = %_CNC.tool_dz;
      %__tmp_tool.Frame.Orient.Type = %_CNC.tool_angles_type;
      %__tmp_tool.Frame.Orient.Angle[0] = %_CNC.tool_phi;
      %__tmp_tool.Frame.Orient.Angle[1] = %_CNC.tool_theta;
      %__tmp_tool.Frame.Orient.Angle[2] = %_CNC.tool_psi;
      %__tmp_tool.Frame.Orient.Angle[3] = 0;
      %__tmp_tool.Radius = #sys_vars.RAD;
    GetTool:
      Arg (ref=Tool, UserType=MXToolType, MinCount=1, MaxCount=1)
    TmpBaseFrame = %__tmp_frame.Pos.x = %_CNC.base_frame_dx;
      %__tmp_frame.Pos.y = %_CNC.base_frame_dy;
      %__tmp_frame.Pos.z = %_CNC.base_frame_dz;
      %__tmp_frame.Orient.Type = %_CNC.base_frame_angles_type;
      %__tmp_frame.Orient.Angle[0] = %_CNC.base_frame_phi;
      %__tmp_frame.Orient.Angle[1] = %_CNC.base_frame_theta;
      %__tmp_frame.Orient.Angle[2] = %_CNC.base_frame_psi;
      %__tmp_frame.Orient.Angle[3] = 0;
    GetBaseFrame:
      Arg (ref=Frame, UserType=MXFrameType, MinCount=1, MaxCount=1)
    GetJoint:
      Arg (ref=Joint, UserType=MXJointAxisType, MinCount=1, MaxCount=1)
    GetAxisTarget:
      Arg (ref=AxisTarget, UserType=MXAxisTargetType, MinCount=1, MaxCount=1)
    GetLatchPoint:
      Arg (ref=ID, DataType=IEC_UINT, MinCount=1, MaxCount=1)
      Arg (ref=Point, UserType=MXPointType, MinCount=1, MaxCount=1)
      Arg (ref=Event, DataType=IEC_BOOL, MinCount=1, MaxCount=1)
    GetPoint:
      Arg (ref=Point, UserType=MXPointType, MinCount=1, MaxCount=1)
    GetPointIntern = %__tmp_point = %POINT_0;
      
      local $i;
      $i=0;
      lbegin(1)
        %__tmp_axis_code[$i] = %_AX.axis_map[$i];
        %__tmp_axis_idx[$i] = %_AX.axis_map_idx[$i];
        $i = $i + 1;
      lend($i < GetIpInt(:300:))     
      %__mx_status =  MXCncAxesToPoint(:%_CNC.adr_trf_data_mx,  \%__tmp_set_pos, \%__tmp_point,   %_CNC.trf_type, %_CNC.angles_type, \%__tmp_axis_code, \%__tmp_axis_idx, GetIpInt(:300:) :);
      if (%__mx_status > 0)
        
        ErrorEx(:"id":10905,"fmt":"4d4d4d","data":(:GetCurLine(::),4,%__mx_status:):);
      endif
    CDCOn:
      Arg (ref=Direction, DataType=INT, MinCount=1, MaxCount=1)
      Arg (ref=CDC, UserType=MXCDCType, MinCount=0, MaxCount=1)
    CDCOff:
      Arg (ref=CDC, UserType=MXCDCType, MinCount=0, MaxCount=1)
    AutoTangOn:
      Arg (ref=Param, UserType=MXAutoTangType, MinCount=0, MaxCount=1)
    AutoTangOff = #next_motion.Command = MPCMD_MX_TANG_AX_OFF;
      PushPacket(::);
    SetM = local $i, $num_item;
      $i = 1;
      $num_item = ListLength(:${*}:);
      lbegin (1)
        #next_motion.Command = MPCMD_SET_M_FCT;
        #next_motion.Data.I4_value = ListItemValue(:${*}, $i:);  
        PushPacket(::);
        $i = $i + 1;
      lend($i <= $num_item)
      DispatchMPList(::); (MinArgs=1, MaxArgs=10)
  SysVars:
    TRF_DATA_MX $TRF_DATA_MX:
      GET = return %_CNC.adr_trf_data_mx; (ReturnType=IEC_UDINT)
```

### Data object Logical/GmcIpUserConfig/gmcipvar (Cnc, version 5.02.1)

#### gmcipvar.cnc
```
CONFIG:
  VARIABLES
```

### Data object Logical/GmcIpUserConfig/gmcipfun (Cnc, version 5.02.1)

#### gmcipfun.cnc
```
CONFIG:
  FUNCTIONS
```

### Data object Logical/GmcIpUserConfig/gmcipfub (Cnc, version 5.02.1)

#### gmcipfub.cnc
```
CONFIG:
  FUBOutputs
  FUBS
  VARIABLES
```

### Data object Logical/GmcIpUserConfig/gmcipubr (Cnc, version 5.02.1)

#### gmcipubr.cnc
```
Root (LangModule=ailgcode, Version=1.0)
```

### Data object Logical/GmcIpUserConfig/gmcipusm (Cnc, version 5.02.1)

#### gmcipusm.cnc
```
Root (LangModule=ailgcode, Version=1.0)
```

### Data object Logical/GmcIpUserConfig/gmcipui (Cnc, version 5.02.1)

#### gmcipui.cnc
```
Root (LangModule=ailgcode, Version=1.0)
```

### Data object Logical/GmcIpUserConfig/gmcipus (Cnc, version 5.02.1)

#### gmcipus.cnc
```
LANGS
```

### Data object Logical/GmcIpUserConfig/gmcipuc (Cnc, version 5.02.1)

#### gmcipuc.cnc
```
CONFIG
```

### Package Logical/gAxis01obj - gAxis01obj

### Data object Logical/gAxis01obj/gAxis01a (Apt)

#### gAxis01a.apt
```
AcoposParameterTable:
  Root Parameters:
    64232 = 51200 (Name=SM_SCALE_STEP)
    64233 = 1000 (Name=SM_SCALE_LOAD_UNITS)
    64234 = 1 (Name=SM_SCALE_LOAD_MOTREV)
    109 = 1024 (Name=SCALE_ENCOD_INCR)
    110 = ncSW_ON (Name=CMD_SIMULATION)
```

### Data object Logical/gAxis01obj/gAxis01i (Ax)

#### gAxis01i.ax
```
InitParameter (Version=5.2.1, NcSwId=Acp10)
  ACP10AXIS_typ:
    dig_in:
      level:
        reference = ncACTIV_HI
        pos_hw_end = ncACTIV_HI
        neg_hw_end = ncACTIV_HI
        trigger1 = ncACTIV_HI
        trigger2 = ncACTIV_HI
    encoder_if:
      parameter:
        count_dir = ncSTANDARD
        scaling:
          load:
            units = 1000
            rev_motor = 1
    limit:
      parameter:
        v_pos = 10000
        v_neg = 10000
        a1_pos = 50000
        a2_pos = 50000
        a1_neg = 50000
        a2_neg = 50000
        t_jolt = 0
        t_in_pos = 0
        pos_sw_end = 2000000000
        neg_sw_end = -2000000000
        ds_warning = 500
        ds_stop = 1000
        a_stop = 1.0e30
        dv_stop = 0
        dv_stop_mode = ncOFF
    controller:
      mode = ncPOSITION
      position:
        kv = 50
        tn = 0
        t_predict = 0.01
        t_total = 0.01
        p_max = 1.0e30
        i_max = 0
      speed:
        kv = 2.0
        tn = 0
        t_filter = 0.0
        isq_filter1:
          type = ncOFF
          a0 = 0.0
          a1 = 0.0
          b0 = 0.0
          b1 = 0.0
          b2 = 0.0
          c0_par_id = 0
          c1_par_id = 0
        isq_filter2:
          type = ncOFF
          a0 = 0.0
          a1 = 0.0
          b0 = 0.0
          b1 = 0.0
          b2 = 0.0
          c0_par_id = 0
          c1_par_id = 0
        isq_filter3:
          type = ncOFF
          a0 = 0.0
          a1 = 0.0
          b0 = 0.0
          b1 = 0.0
          b2 = 0.0
          c0_par_id = 0
          c1_par_id = 0
      uf:
        type = ncLINEAR + ncCORRECTION
        auto_config = ncMOTOR_PAR
        u0 = 0
        un = 0
        fn = 50.0
        k_f_slip = 0
      ff:
        torque_load = 0.0
        torque_pos = 0.0
        torque_neg = 0.0
        kv_torque = 0.0
        inertia = 0.0
        t_filter_a = 0.0
    move:
      stop:
        parameter[0]:
          decel_ramp = ncA_LIMIT
          controller = ncON
        parameter[1]:
          decel_ramp = ncA_LIMIT
          controller = ncON
        parameter[2]:
          decel_ramp = ncA_LIMIT
          controller = ncON
        parameter[3]:
          decel_ramp = ncA_LIMIT
          controller = ncON
        quickstop:
          decel_ramp = ncA_LIMIT
          t_jolt = 0
        drive_error:
          decel_ramp = ncA_LIMIT
      homing:
        parameter:
          s = 0
          v_switch = 5000
          v_trigger = 500
          a = 50000
          mode = ncDIRECT
          edge_sw = ncPOSITIVE
          start_dir = ncPOSITIVE
          trigg_dir = ncPOSITIVE
          ref_pulse = ncOFF
          fix_dir = ncOFF
          tr_s_block = 0
          torque_lim = 0
          ds_block = 0
          ds_stop = 0
      basis:
        parameter:
          v_pos = 5000
          v_neg = 5000
          a1_pos = 50000
          a2_pos = 50000
          a1_neg = 50000
          a2_neg = 50000
    message:
      text:
        parameter:
          format = ncBREAK
          columns = 80
          data_modul = acp10etxen
```

### Program Logical/Program (ANSIC)

#### Main.c - Init, cyclic, exit code
```c
#include <bur/plctypes.h>

#ifdef _DEFAULT_INCLUDES
	#include <AsDefault.h>
#endif

void _INIT ProgramInit(void)
{

}

void _CYCLIC ProgramCyclic(void)
{
	doorSM.state = stateMachine.state;
	DoorStateMachine(&doorSM);

	stateMachine.enable = 1;
	stateMachine.setSpeed = doorSM.speed;
	DriveStateMachine(&stateMachine);

	ledSM.state = doorSM.doorState;
	LedStateMachine(&ledSM);

}

void _EXIT ProgramExit(void)
{

}
```

### Library Logical/Library (ANSIC)

#### Types.typ - Exported data types
```iecst
TYPE
	DoorStates :
		(
		ST_INIT,
		ST_UNKNOWN,
		ST_OPEN,
		ST_CLOSE,
		ST_ACC_POS,
		ST_ACC_NEG,
		ST_POS,
		ST_NEG,
		ST_DEC_POS,
		ST_DEC_NEG
		);
END_TYPE
```

#### Library.fun - Exported functions and function blocks
```iecst
{REDUND_ERROR} FUNCTION_BLOCK DriveStateMachine (*TODO: Add your comment here*) (*$GROUP=User,$CAT=User,$GROUPICON=User.png,$CATICON=User.png*)
	VAR_INPUT
		state : {REDUND_UNREPLICABLE} UINT;
		enable : {REDUND_UNREPLICABLE} BOOL := 0;
		setSpeed : {REDUND_UNREPLICABLE} INT;
	END_VAR
	VAR_OUTPUT
		command : {REDUND_UNREPLICABLE} UINT;
		speed : {REDUND_UNREPLICABLE} INT;
	END_VAR
	VAR
		step : {REDUND_UNREPLICABLE} USINT;
	END_VAR
END_FUNCTION_BLOCK

{REDUND_ERROR} {REDUND_UNREPLICABLE} FUNCTION_BLOCK DoorStateMachine (*TODO: Add your comment here*) (*$GROUP=User,$CAT=User,$GROUPICON=User.png,$CATICON=User.png*)
	VAR_INPUT
		state : {REDUND_UNREPLICABLE} UINT;
		sw1 : {REDUND_UNREPLICABLE} BOOL;
		sw2 : {REDUND_UNREPLICABLE} BOOL;
		sw3 : {REDUND_UNREPLICABLE} BOOL;
		sw4 : {REDUND_UNREPLICABLE} BOOL;
		direction : {REDUND_UNREPLICABLE} BOOL;
	END_VAR
	VAR_OUTPUT
		speed : {REDUND_UNREPLICABLE} INT;
	END_VAR
	VAR
		doorState : {REDUND_UNREPLICABLE} DoorStates;
		sw1old : {REDUND_UNREPLICABLE} BOOL;
		sw4old : {REDUND_UNREPLICABLE} BOOL;
		sw3old : {REDUND_UNREPLICABLE} BOOL;
		sw2old : {REDUND_UNREPLICABLE} BOOL;
	END_VAR
END_FUNCTION_BLOCK

{REDUND_ERROR} {REDUND_UNREPLICABLE} FUNCTION_BLOCK LedStateMachine (*TODO: Add your comment here*) (*$GROUP=User,$CAT=User,$GROUPICON=User.png,$CATICON=User.png*)
	VAR_INPUT
		state : {REDUND_UNREPLICABLE} UINT;
	END_VAR
	VAR_OUTPUT
		led1 : {REDUND_UNREPLICABLE} BOOL;
		led2 : {REDUND_UNREPLICABLE} BOOL;
		led3 : {REDUND_UNREPLICABLE} BOOL;
		led4 : {REDUND_UNREPLICABLE} BOOL;
		timer : {REDUND_UNREPLICABLE} INT;
	END_VAR
END_FUNCTION_BLOCK
```

#### DriveStateMachine.c
```c
#include <bur/plctypes.h>
#ifdef __cplusplus
	extern "C"
	{
#endif
	#include "Library.h"
#ifdef __cplusplus
	};
#endif
/* TODO: Add your comment here */
#define CMD_SHUTDOWN 0x06
#define CMD_SWITCH_ON 0x07
#define CMD_ENABLE 0x0F
#define CMD_FAULT_RESET 0x80

#define STATE_MASK 0x6F
#define STATE_READY_TO_SWITCH_ON 0x21
#define STATE_SWITCHED_ON 0x23
#define STATE_OP_ENABLED 0x27
#define STATE_FAULT_BIT 0x08

void DriveStateMachine(struct DriveStateMachine* inst)
{
	UINT st = inst->state & STATE_MASK;

	switch (inst->step){
		case 0:
			inst->speed = 0;
			inst->command = (inst->state & STATE_FAULT_BIT) ? CMD_FAULT_RESET : CMD_SHUTDOWN;
			if (inst->enable && st == STATE_READY_TO_SWITCH_ON)
				inst->step = 1;
			break;
		case 1:
			inst->speed = 0;
			inst->command = CMD_SWITCH_ON;
			if (!inst->enable) inst->step = 0;
			else if (st == STATE_SWITCHED_ON) inst->step = 2;
		case 2:
			inst->command = CMD_ENABLE;
			inst->speed = inst->setSpeed;
			if (!inst->enable || (inst->state & STATE_FAULT_BIT))
				inst->step = 0;
			break;
	}

}
```

#### DoorStateMachine.c
```c
#include <bur/plctypes.h>
#ifdef __cplusplus
	extern "C"
	{
#endif
	#include "Library.h"
#ifdef __cplusplus
	};
#endif
/* TODO: Add your comment here */
#define V_FAST 600
#define V_SLOW 150
#define CMD_CLOSE 1
#define DRV_OP_ENABLED 0x27

void DoorStateMachine(struct DoorStateMachine* inst)
{
	INT v = 0;
	BOOL closeCMD = (inst->direction == CMD_CLOSE);

	if ((inst->state & 0x6F) != DRV_OP_ENABLED){
		inst->doorState = ST_INIT;
	}
	BOOL sw1_ch = (inst->sw1 != inst->sw1old);
	BOOL sw2_ch = (inst->sw2 != inst->sw2old);
	BOOL sw3_ch = (inst->sw3 != inst->sw3old);
	BOOL sw4_ch = (inst->sw4 != inst->sw4old);

	inst->sw1old = inst->sw1;
	inst->sw2old = inst->sw2;
	inst->sw3old = inst->sw3;
	inst->sw4old = inst->sw4;

	switch (inst->doorState){
		case ST_INIT:
			v = 0;
			if ((inst->state & 0x6F) == DRV_OP_ENABLED){
				inst->doorState = ST_UNKNOWN;
			}
			break;

		case ST_UNKNOWN:
			if (closeCMD) {
				v = V_SLOW;
				if (sw4_ch){
					inst->doorState = ST_CLOSE;
				}}
			else {
				v = -V_SLOW;
				if (sw1_ch){
					inst->doorState = ST_OPEN;
				}
			}
			break;

		case ST_OPEN:
			v = 0;
			if (closeCMD && sw1_ch){
				inst->doorState = ST_ACC_POS;
			}
			break;

		case ST_ACC_POS:
			v = V_SLOW;
			if (sw2_ch) {
				inst->doorState = ST_POS;
			}
			else if (!closeCMD){
				inst->doorState = ST_DEC_NEG;
			}
			break;

		case ST_POS:
			v = V_FAST;
			if (sw3_ch) {
				inst->doorState = ST_DEC_POS;
			}
			else if (!closeCMD){
				inst->doorState = ST_NEG;
			}
			break;

		case ST_DEC_POS:
			v = V_SLOW;
			if (sw4_ch) {
				inst->doorState = ST_CLOSE;
			}
			else if (!closeCMD){
				inst->doorState = ST_ACC_NEG;
			}
			break;

		case ST_CLOSE:
			v = 0;
			if (!closeCMD && sw4_ch){
				inst->doorState = ST_ACC_NEG;
			}
			break;

		case ST_ACC_NEG:
			v = -V_SLOW;
			if (sw3_ch) {
				inst->doorState = ST_NEG;
			}
			else if (closeCMD){
				inst->doorState = ST_DEC_POS;
			}
			break;

		case ST_NEG:
			v = -V_FAST;
			if (sw2_ch) {
				inst->doorState = ST_DEC_NEG;
			}
			else if (closeCMD){
				inst->doorState = ST_POS;
			}
			break;

		case ST_DEC_NEG:
			v = -V_SLOW;
			if (sw1_ch) {
				inst->doorState = ST_OPEN;
			}
			else if (closeCMD){
				inst->doorState = ST_ACC_POS;
			}
			break;
	}
	inst->speed = v;
}
```

#### LedStateMachine.c
```c
#include <bur/plctypes.h>
#ifdef __cplusplus
	extern "C"
	{
#endif
#include "Library.h"
#ifdef __cplusplus
	};
#endif
/* TODO: Add your comment here */
#define CYCLE_MS 10

static void setLeds(struct LedStateMachine* inst, BOOL a, BOOL b,BOOL c,BOOL d){
	inst->led1 = a;
	inst->led2 = b;
	inst->led3 = c;
	inst->led4 = d;
}

void LedStateMachine(struct LedStateMachine* inst)
{
	BOOL blink;

	switch (inst->state){
		case ST_UNKNOWN:
			inst->timer +=CYCLE_MS;
			if (inst->timer >= 1000) inst->timer = 0;
			blink = (inst->timer < 500);
			setLeds(inst, blink, blink, blink, blink);
			return;

		case ST_ACC_POS: case ST_DEC_NEG: setLeds(inst, 1,0,0,0); break;
		case ST_POS: case ST_NEG: setLeds(inst, 1,1,0,0); break;
		case ST_DEC_POS: case ST_ACC_NEG: setLeds(inst, 1,1,1,0); break;
		case ST_CLOSE: setLeds(inst, 1,1,1,1); break;
		default: setLeds(inst, 0,0,0,0); break;
	}
	inst->timer = 0;
}
```
